Fanuc KAREL source: KC00032.KL

PROGRAM KC00032
%NOLOCKGROUP
%ENVIRONMENT BYNAM
VAR
  I: INTEGER
  J: INTEGER
  K: INTEGER
  R: REAL
  B: BOOLEAN
  S: STRING[80]
  T: STRING[80]
  P: PATH
  Q: PATH
  AI: ARRAY[8] OF INTEGER
  AB: ARRAY[244] OF BYTE
  SA: ARRAY[8] OF STRING[80]
BEGIN
  PROG_LIST(S,I,J,K,SA,I,J)
END KC00032
